// TwinCAT 3 PLC project MainControl
// ProgramVersion: 3.1.4024.0
// libraries:
//   JS_MC_REF, * (Jenny Science AG)
//   Tc2_EtherCAT, * (Beckhoff Automation GmbH)
//   Tc2_MC2, * (Beckhoff Automation GmbH)
//   Tc2_NCI, * (Beckhoff Automation GmbH)
//   Tc2_PlcInterpolation, * (Beckhoff Automation GmbH)
//   Tc2_Standard, * (Beckhoff Automation GmbH)
//   Tc2_System, * (Beckhoff Automation GmbH)
//   Tc2_Utilities, * (Beckhoff Automation GmbH)
//   Tc3_Module, * (Beckhoff Automation GmbH)
// project tree:
//   DUTs/ MFuncs.TcDUT, T_StringQueue.TcDUT
//   GVLs/ ExtPort.TcGVL, HMIVar.TcGVL, PYADSPort.TcGVL, UserVar.TcGVL
//   / PlcTask.TcTTO
//   POUs/FB/ FB_BackendManager.TcPOU, FB_ExtMessage.TcPOU, FB_HMITask.TcPOU, FB_JSReference.TcPOU, FB_Jog.TcPOU, FB_McodeMonitor.TcPOU, FB_MotorPower.TcPOU, FB_MotorReset.TcPOU, FB_RParamInit.TcPOU, FB_TimeCalculator.TcPOU
//   POUs/FB/Keyence/ FB_LJ_S8000Capture.TcPOU
//   POUs/FB/MicroFab/ FB_PulseInterval.TcPOU
//   POUs/FB/Nordson/ FB_ReadPressure.TcPOU, FB_WritePressure.TcPOU
//   POUs/function/ f_Contains_INT.TcPOU, f_MakeAbsPath.TcPOU, f_QueuePop.TcPOU, f_QueuePush.TcPOU, f_Queue_ToString.TcPOU
//   POUs/ MotorControl.TcPOU
// real-time tasks:
//   TASK PlcTask: cycle T#10ms, priority 20, ADS port 350
// motion (NC):
//   TASK NC-Task 1 SAF: cycle T#1ms, priority 4, ADS port 501
//   TASK NC-Task 1 SVB: cycle T#10ms, priority 8, ADS port 511
//   AXIS Axis 1 (id 1)
//     Velo: SlowManual=5, FastManual=30, Maximum=4500
//     OtherSettings: AllowMotionCmdToSlave=true
//     encoder EncType=19
//       EncPara: ScaleFactorNumerator=0.001, MaxCount=#xffffffff
//     drive DrvType=16
//       DrvPara: MaxCount=#xffffffff, DriveControlDWord=#x00020100
//         Analog: VeloReferenz=4500, VeloScale=125, AccScale=0.02, TorqueSetpointScale=10, ScaleFactorActTorque=0.1
//         TimeComp: TaskDelayCycles=1
//     controller CtrType=9
//       CtrPara: PriorControlFactor=1
//         Observer: BandWidth=20
//   AXIS Axis 2 (id 2)
//     Velo: SlowManual=5, FastManual=30, Maximum=4500
//     OtherSettings: AllowMotionCmdToSlave=true
//     encoder EncType=19
//       EncPara: ScaleFactorNumerator=0.001, MaxCount=#xffffffff
//     drive DrvType=16
//       DrvPara: MaxCount=#xffffffff, DriveControlDWord=#x00020100
//         Analog: VeloReferenz=4500, VeloScale=125, AccScale=0.02, TorqueSetpointScale=10, ScaleFactorActTorque=0.1
//         TimeComp: TaskDelayCycles=1
//     controller CtrType=9
//       CtrPara: PriorControlFactor=1
//         PID: PosKp=0
//         Observer: BandWidth=20
//   AXIS Axis 3 (id 3)
//     Velo: SlowManual=5, FastManual=30, Maximum=4500
//     OtherSettings: AllowMotionCmdToSlave=true
//     encoder EncType=19
//       EncPara: ScaleFactorNumerator=0.001, MaxCount=#xffffffff
//     drive DrvType=16
//       DrvPara: MaxCount=#xffffffff, DriveControlDWord=#x00020100
//         Analog: VeloReferenz=4500, VeloScale=125, AccScale=0.02, TorqueSetpointScale=10, ScaleFactorActTorque=0.1
//         TimeComp: TaskDelayCycles=1
//     controller CtrType=9
//       CtrPara: PriorControlFactor=1
//         Observer: BandWidth=20
//   AXIS Axis 4 (id 4)
//     Velo: SlowManual=1, FastManual=5
//     OtherSettings: AllowMotionCmdToSlave=true
//     encoder EncType=19
//       EncPara: MaxCount=#xffffffff
//     drive DrvType=16
//       DrvPara: MaxCount=#xffffffff, DriveControlDWord=#x00020000
//         Analog: TorqueSetpointScale=10, ScaleFactorActTorque=0.1
//         TimeComp: TaskDelayCycles=1
//     controller CtrType=1
//       CtrPara: PriorControlFactor=1
//         Observer: BandWidth=20
// I/O:
//   DEVICE Device 2 (EtherCAT), AmsNetId 192.168.0.2.3.1
//     Drive 1 (Xvi) [XENAX Xvi 75V8S]
//     Drive 2 (Xvi) [XENAX Xvi 75V8S]
//     Drive 3 (Xvi) [XENAX Xvi 75V8S]
//     Drive 12 (Ezi-SERVO2 EtherCAT) [Ezi-SERVO2 EtherCAT]
//     Term 4 (EK1100) [EK1100 EtherCAT Coupler (2A E-Bus)]
//       Term 5 (EL1008) [EL1008 8Ch. Dig. Input 24V, 3ms]
//       Term 17 (EL2008) [EL2008 8Ch. Dig. Output 24V, 0.5A]
//       Term 6 (EL9185) [EL9185 Potential Connection, 4 x 24-230V]
//       Term 7 (EL9505) [EL9505 Power supply terminal 5V]
//       Term 10 (EL2124) [EL2124 4Ch. Dig. Output 5V, 20mA]
//       Term 11 (EL2634) [EL2634 4Ch. Relay Output, NO (250V AC / 30V DC)]
//       Term 9 (EL9011) [EL9011 End Terminal]
//     Box 8 (LJ-S_CB-NEC Series) [LJ-S_CB-NEC Series]
//       modules: Module 1 (Result Data 128Byte), Module 2 (Parameter 128Byte)
// variable links:
//   NC-Task 1 SAF/Axes/Axis 1 <-> Device 2 (EtherCAT)/Drive 1 (Xvi)
//     Drive/Inputs/In/nDataIn1 <-> 1. TxPDO CSP/Following Error Actual Value
//     Drive/Inputs/In/nState1 <-> 1. TxPDO CSP/Statusword
//     Drive/Inputs/In/nState2 <-> 1. TxPDO CSP/Statusword @bit 8
//     Drive/Inputs/In/nState4 @bit 1 <-> WcState/InputToggle
//     Drive/Inputs/In/nState4 <-> WcState/WcState
//     Drive/Outputs/Out/nCtrl1 <-> 1. RxPDO CSP/Controlword
//     Drive/Outputs/Out/nCtrl2 <-> 1. RxPDO CSP/Controlword @bit 8
//     Drive/Outputs/Out/nDataOut1 <-> 1. RxPDO CSP/Target Position
//     Drive/Outputs/Out/nDataOut2 <-> 4. RxPDO CSP FeedForward/Target Velocity
//     Drive/Outputs/Out/nDataOut3[0] <-> 4. RxPDO CSP FeedForward/Torque Offset
//     Enc/Inputs/In/nDataIn1 <-> 1. TxPDO CSP/Position Actual Value
//     Enc/Inputs/In/nState4 @bit 1 <-> WcState/InputToggle
//     Enc/Inputs/In/nState4 <-> WcState/WcState
//   NC-Task 1 SAF/Axes/Axis 2 <-> Device 2 (EtherCAT)/Drive 2 (Xvi)
//     Drive/Inputs/In/nDataIn1 <-> 1. TxPDO CSP/Following Error Actual Value
//     Drive/Inputs/In/nState1 <-> 1. TxPDO CSP/Statusword
//     Drive/Inputs/In/nState2 <-> 1. TxPDO CSP/Statusword @bit 8
//     Drive/Inputs/In/nState4 @bit 1 <-> WcState/InputToggle
//     Drive/Inputs/In/nState4 <-> WcState/WcState
//     Drive/Outputs/Out/nCtrl1 <-> 1. RxPDO CSP/Controlword
//     Drive/Outputs/Out/nCtrl2 <-> 1. RxPDO CSP/Controlword @bit 8
//     Drive/Outputs/Out/nDataOut1 <-> 1. RxPDO CSP/Target Position
//     Drive/Outputs/Out/nDataOut2 <-> 4. RxPDO CSP FeedForward/Target Velocity
//     Drive/Outputs/Out/nDataOut3[0] <-> 4. RxPDO CSP FeedForward/Torque Offset
//     Enc/Inputs/In/nDataIn1 <-> 1. TxPDO CSP/Position Actual Value
//     Enc/Inputs/In/nState4 @bit 1 <-> WcState/InputToggle
//     Enc/Inputs/In/nState4 <-> WcState/WcState
//   NC-Task 1 SAF/Axes/Axis 3 <-> Device 2 (EtherCAT)/Drive 3 (Xvi)
//     Drive/Inputs/In/nDataIn1 <-> 1. TxPDO CSP/Following Error Actual Value
//     Drive/Inputs/In/nState1 <-> 1. TxPDO CSP/Statusword
//     Drive/Inputs/In/nState2 <-> 1. TxPDO CSP/Statusword @bit 8
//     Drive/Inputs/In/nState4 @bit 1 <-> WcState/InputToggle
//     Drive/Inputs/In/nState4 <-> WcState/WcState
//     Drive/Outputs/Out/nCtrl1 <-> 1. RxPDO CSP/Controlword
//     Drive/Outputs/Out/nCtrl2 <-> 1. RxPDO CSP/Controlword @bit 8
//     Drive/Outputs/Out/nDataOut1 <-> 1. RxPDO CSP/Target Position
//     Drive/Outputs/Out/nDataOut2 <-> 4. RxPDO CSP FeedForward/Target Velocity
//     Drive/Outputs/Out/nDataOut3[0] <-> 4. RxPDO CSP FeedForward/Torque Offset
//     Enc/Inputs/In/nDataIn1 <-> 1. TxPDO CSP/Position Actual Value
//     Enc/Inputs/In/nState4 @bit 1 <-> WcState/InputToggle
//     Enc/Inputs/In/nState4 <-> WcState/WcState
//   NC-Task 1 SAF/Axes/Axis 4 <-> Device 2 (EtherCAT)/Drive 12 (Ezi-SERVO2 EtherCAT)
//     Drive/Inputs/In/nDcOutputTime <-> InfoData/DcOutputShift
//     Drive/Inputs/In/nState1 <-> CSP Inputs/Status Word
//     Drive/Inputs/In/nState2 <-> CSP Inputs/Status Word @bit 8
//     Drive/Inputs/In/nState4 @bit 1 <-> WcState/InputToggle
//     Drive/Inputs/In/nState4 <-> WcState/WcState
//     Drive/Outputs/Out/nCtrl1 <-> CSP Outputs/Control Word
//     Drive/Outputs/Out/nCtrl2 <-> CSP Outputs/Control Word @bit 8
//     Drive/Outputs/Out/nDataOut1 <-> CSP Outputs/Target Position
//     Enc/Inputs/In/nDataIn1 <-> CSP Inputs/Position Actual Value
//     Enc/Inputs/In/nDataIn3 <-> CSP Inputs/Touch probe 1 positive value
//     Enc/Inputs/In/nDataIn5 <-> CSP Inputs/Touch probe 2 positive value
//     Enc/Inputs/In/nDcInputTime <-> InfoData/DcInputShift
//     Enc/Inputs/In/nState4 @bit 1 <-> WcState/InputToggle
//     Enc/Inputs/In/nState4 <-> WcState/WcState
//     Enc/Inputs/In/nState5 <-> CSP Inputs/Touch probe status
//     Enc/Inputs/In/nState6 <-> CSP Inputs/Touch probe status @bit 8
//     Enc/Outputs/Out/nCtrl5 <-> CSP Outputs/Touch probe function
//     Enc/Outputs/Out/nCtrl6 <-> CSP Outputs/Touch probe function @bit 8
//   MainControl/MainControl Instance <-> Device 2 (EtherCAT)/Box 8 (LJ-S_CB-NEC Series)
//     PlcTask Inputs/ExtPort.LJ_S8000_bBusy <-> StatusBit/BUSY
//     PlcTask Inputs/ExtPort.LJ_S8000_bReady <-> StatusBit/READY
//     PlcTask Inputs/ExtPort.LJ_S8000_bTRG_ack <-> StatusBit/TRG_ack
//     PlcTask Outputs/ExtPort.LJ_S8000_bTRG <-> ControlBit/TRG
//   MainControl/MainControl Instance <-> Device 2 (EtherCAT)/Drive 1 (Xvi)
//     PlcTask Inputs/MotorControl.fb_JSReference.JS_MC_X.stSlaveAmsAddr <-> InfoData/AdsAddr
//   MainControl/MainControl Instance <-> Device 2 (EtherCAT)/Drive 2 (Xvi)
//     PlcTask Inputs/MotorControl.fb_JSReference.JS_MC_Y.stSlaveAmsAddr <-> InfoData/AdsAddr
//   MainControl/MainControl Instance <-> Device 2 (EtherCAT)/Drive 3 (Xvi)
//     PlcTask Inputs/MotorControl.fb_JSReference.JS_MC_Z.stSlaveAmsAddr <-> InfoData/AdsAddr
//   MainControl/MainControl Instance <-> Device 2 (EtherCAT)/Term 4 (EK1100)/Term 10 (EL2124)
//     PlcTask Outputs/ExtPort.EL2124_OUT[0] <-> Channel 1/Output
//   MainControl/MainControl Instance <-> Device 2 (EtherCAT)/Term 4 (EK1100)/Term 11 (EL2634)
//     PlcTask Outputs/ExtPort.EL2634_OUT[0] <-> Channel 1/Output
//   MainControl/MainControl Instance <-> Device 2 (EtherCAT)/Term 4 (EK1100)/Term 5 (EL1008)
//     PlcTask Inputs/ExtPort.EL1008_IN[0] <-> Channel 1/Input
//     PlcTask Inputs/ExtPort.EL1008_IN[1] <-> Channel 2/Input
//   MainControl/MainControl Instance <-> NC-Task 1 SAF/Axes/Axis 1
//     PlcTask Inputs/MotorControl.motX.NcToPlc <-> Outputs/ToPlc
//     PlcTask Outputs/MotorControl.motX.PlcToNc <-> Inputs/FromPlc
//   MainControl/MainControl Instance <-> NC-Task 1 SAF/Axes/Axis 2
//     PlcTask Inputs/MotorControl.motY.NcToPlc <-> Outputs/ToPlc
//     PlcTask Outputs/MotorControl.motY.PlcToNc <-> Inputs/FromPlc
//   MainControl/MainControl Instance <-> NC-Task 1 SAF/Axes/Axis 3
//     PlcTask Inputs/MotorControl.motZ.NcToPlc <-> Outputs/ToPlc
//     PlcTask Outputs/MotorControl.motZ.PlcToNc <-> Inputs/FromPlc
//   MainControl/MainControl Instance <-> NC-Task 1 SAF/Axes/Axis 4
//     PlcTask Inputs/MotorControl.motQ1.NcToPlc <-> Outputs/ToPlc
//     PlcTask Outputs/MotorControl.motQ1.PlcToNc <-> Inputs/FromPlc
//   MainControl/MainControl Instance <-> NC-Task 1 SAF/Channel 2
//     PlcTask Inputs/MotorControl.inst_NcToPlc_NCI <-> Outputs/ToPlc
//     PlcTask Outputs/MotorControl.inst_PlcToNc_NCI <-> Inputs/FromPlc

CONFIGURATION MainControl
    RESOURCE PLC ON TwinCAT3
        TASK PlcTask(INTERVAL := T#10ms, PRIORITY := 20);
        PROGRAM MotorControl WITH PlcTask : MotorControl;
    END_RESOURCE
END_CONFIGURATION

// ---- DUTs/MFuncs.TcDUT
TYPE MFuncs :
//	M: 0 ~ 159
//	NOT TO USE THESE M-FUNCTIONS
//  2	(Program end)
//	17	(End of subprogram)
//	30	(Program end with delection of all fast M functions)
(
	M_NordsonExtOn		:=	10,
	M_NordsonExtOff 	:=	11,

	M_MicrofabExtOn		:=	20,
	M_MicrofabExtOff	:=	21,
	
	M_LJ_S8000TRG		:=	50,
	
	
	M_NordsonPresTRG100	:=	100,
	M_NordsonPresTRG101	:=	101,
	M_NordsonPresTRG102	:=	102,
	M_NordsonPresTRG103	:=	103,
	M_NordsonPresTRG104	:=	104,
	M_NordsonPresTRG105	:=	105,
	M_NordsonPresTRG106	:=	106,
	M_NordsonPresTRG107	:=	107,
	M_NordsonPresTRG108	:=	108,
	M_NordsonPresTRG109	:=	109,
	
	M_MicrofabIntTRG110 :=	110,
	M_MicrofabIntTRG111 :=	111,
	M_MicrofabIntTRG112 :=	112,
	
	
	M_RHskTRG			:=	150
	
);
END_TYPE

// ---- DUTs/T_StringQueue.TcDUT
TYPE T_StringQueue :
STRUCT
    Buffer : ARRAY[0..19] OF STRING(255); // 큐 크기 20
    Head   : INT	:=	0;  // Pop 위치
    Tail   : INT	:=	0;  // Push 위치
    Count  : INT	:=	0;  // 현재 개수
END_STRUCT
END_TYPE

// ---- GVLs/ExtPort.TcGVL
{attribute 'qualified_only'}
VAR_GLOBAL
	// ExtPort.EL2124_OUT[0]	:	MicroFab Ext 1
	EL2124_OUT	AT%Q*	:	ARRAY[0..3]	OF	BOOL;
	
	// ExtPort.EL2634_OUT[0]	:	Nordson Ext 1
	EL2634_OUT	AT%Q*	:	ARRAY[0..3]	OF	BOOL;
	
	LJ_S8000_bBusy		AT%I*	:	BOOL;
	LJ_S8000_bTRG_ack	AT%I*	:	BOOL;
	LJ_S8000_bReady		AT%I*	:	BOOL;
	LJ_S8000_bTRG		AT%Q*	:	BOOL;
	
	EL1008_IN	AT%I*	:	ARRAY[0..7]	OF	BOOL;
END_VAR

// ---- GVLs/HMIVar.TcGVL
{attribute 'qualified_only'}
VAR_GLOBAL
	
	sActPosX	:	STRING(32)	:=	'0.000';
	sActPosY	:	STRING(32)	:=	'0.000';
	sActPosZ	:	STRING(32)	:=	'0.000';
	
	sActVelX	:	STRING(32)	:=	'0.000';
	sActVelY	:	STRING(32)	:=	'0.000';
	sActVelZ	:	STRING(32)	:=	'0.000';
	
	sActAccX	:	STRING(32)	:=	'0.000';
	sActAccY	:	STRING(32)	:=	'0.000';
	sActAccZ	:	STRING(32)	:=	'0.000';
	
	sSetPosX	:	STRING(32)	:=	'0.000';
	sSetPosY	:	STRING(32)	:=	'0.000';
	sSetPosZ	:	STRING(32)	:=	'0.000';
	
	sSetVelX	:	STRING(32)	:=	'0.000';
	sSetVelY	:	STRING(32)	:=	'0.000';
	sSetVelZ	:	STRING(32)	:=	'0.000';
	
	sSetAccX	:	STRING(32)	:=	'0.000';
	sSetAccY	:	STRING(32)	:=	'0.000';
	sSetAccZ	:	STRING(32)	:=	'0.000';
	
	
	EstimatedTime		:	STRING(32)	:=	'0.000s';
	
	
	bNaviActive	:	BOOL	:=	TRUE;
	
	CodeName	:	STRING(255);
	
	GCodeQueueString:	STRING(8192):=	'';
	
	NordsonPressure			:	STRING	:=	'0';
	
	
	I_ForceActX		AT%I*	:	DINT;
	I_ForceActY		AT%I*	:	DINT;
	I_ForceActZ		AT%I*	:	DINT;
	
	
	RunningGCodeLine	:	STRING(1024)	:=	'';
	
	CurrBlockNumSTR		:	STRING	:=	'-';
	
	
	
END_VAR

// ---- GVLs/PYADSPort.TcGVL
{attribute 'qualified_only'}
VAR_GLOBAL
	// Nordson
	bNordWriteReq	:	BOOL	:=	FALSE;
	bNordWriteErr	:	BOOL	:=	FALSE;
	bNordReadReq	:	BOOL	:=	FALSE;
	bNordReadErr	:	BOOL	:=	FALSE;
	nNordPress		:	REAL	:=	0.0;
	
	
	bHeartbeat		:	BOOL	:=	FALSE;
	dtHeartbeatTime	:	DT;
	
	bEstTimeReq		:	BOOL	:=	FALSE;
	bEstTimeErr		:	BOOL	:=	FALSE;
	nEstTime		:	REAL	:=	0.0;	
	
END_VAR

// ---- GVLs/UserVar.TcGVL
{attribute 'qualified_only'}
VAR_GLOBAL
	
	RunningGCodeName:	STRING(255)	:=	'';
//	QueuedGCodeName	:	STRING(255)	:=	'';
	GCodeNameQueue	:	T_StringQueue;
	
	ContinueGCode	:	BOOL	:=	TRUE;
	
	SingleGCodeMode	:	BOOL	:=	FALSE;
	SingleGCodeTRG	:	BOOL	:=	FALSE;
	
	// 0: OFF, 1: JOG, 2: GCODE
	OpMode	:	UDINT	:=	0;
	
	// 0: Nothing, +1: +, +2: ++, -1: -, -2: --
	// +-3: ManualVel 
	JogButtonX	:	INT	:=	0;
	JogButtonY	:	INT	:=	0;
	JogButtonZ	:	INT	:=	0;
//	JogVel		:	LREAL	:=	30.0;
	
	JogMovePos	:	BOOL	:=	FALSE;
	JogTargX	:	STRING	:=	'100.0';
	JogTargY	:	STRING	:=	'260.0';
	JogTargZ	:	STRING	:=	'60.0';
	JogTargVel	:	STRING	:=	'1800'; // Feedrate (mm/min)
	
	JogPowerX	:	BOOL	:=	TRUE;
	JogPowerY	:	BOOL	:=	TRUE;
	JogPowerZ	:	BOOL	:=	TRUE;
	
	NordsonReadPressureBtn	:	BOOL	:=	FALSE;
	NordsonWritePressureBtn	:	BOOL	:=	FALSE;
	NordsonPressureActive	:	BOOL	:=	TRUE;
	
	LJ_S8000CaptureBtn		:	BOOL	:=	FALSE;
	LJ_S8000CaptureActive	:	BOOL	:=	TRUE;
	
	GCodeBasePath	:	STRING(255)	:=	'C:\\Users\\Administrator\\Desktop\\GCodes';

	// 0: Don't input HMIVar.CodeName into execution
	// 1: HMIVar.CodeName into QueuedGCodeName
	// 2: HMIVar.CodeName into GCodeName LIST
	Auto_CodeType	:	INT	:=	1;
	
	R_Params		:	ARRAY[0..12] OF INT	:=
						[100, 101, 102, 103, 104, 105, 106, 107, 108, 109,
						 110, 111, 112];
	
	R_InitVal		:	LREAL	:=	-1.0;
	
	bBackendStarted	:	BOOL	:=	FALSE;
	
	//	gDtFromPy : DT;      // Python이 써주는 시간(권장: UTC epoch seconds로 써서 DT에 저장)
//    gPlcNowDt : DT;      // PLC 로컬 현재시간을 DT로 변환해 저장(옵션)
    gDiffSec  : LINT;    // (PLC - Python) 차이[초]
    gInSync   : BOOL	:=	TRUE;    // 동기 여부
	gPlcStr: STRING(24);
    gPyStr    : STRING(24);
	
	bClearQueue	:	BOOL	:=	FALSE;
	
	
	bESTOP		:	BOOL	:=	FALSE;
	bRESET		:	BOOL	:=	FALSE;
	
	
	bSingleBlockMode	:	BOOL	:=	FALSE;
	
	bNordsonFoot	:	BOOL	:=	FALSE;
	
	CurrBlockNum		:	UDINT	:=	0;
	// Optional Axis 4. Non-retained; all motion permissions default OFF.
	Q1Commissioned : BOOL := FALSE; // Operator confirmation; NOT a safety function
	Q1Enable : BOOL := FALSE;
	Q1UseInGCode : BOOL := FALSE; // Sampled in state 200, held for whole queue run
	Q1Reset : BOOL := FALSE; // Rising edge, idle only
	Q1JogButton : INT := 0; // -1 / 0 / +1 only
	Q1JogVelocity : LREAL := 0.0; // NC units/second; validate before setting
END_VAR

// ---- POUs/MotorControl.TcPOU
PROGRAM MotorControl
VAR
	motX	:	AXIS_REF;
	motY	:	AXIS_REF;
	motZ	:	AXIS_REF;
	
	inst_NcToPlc_NCI	AT %I*	:	NCTOPLC_NCICHANNEL_REF;
	inst_PlcToNc_NCI	AT %Q*	:	PLCTONC_NCICHANNEL_REF;
	
	fb_JSReference	:	FB_JSReference;
	fb_MotorPower	:	FB_MotorPower;
	fb_MotorReset	:	FB_MotorReset;
	
	fb_McodeMonitor	:	FB_McodeMonitor;
	fb_RParamInit	:	FB_RParamInit;
	fb_Backend		:	FB_BackendManager;
	
	bPowered	:	BOOL;
	bMotorReset	:	BOOL;
	bError		:	BOOL;
	bBusy		:	BOOL;
	
	bOpMcodeMonitor	:	BOOL	:=	FALSE;
	
	nMotorControlState	:	UDINT	:= 0;
	nInterpreterState	:	UDINT	:= 0;
	nErrorState			:	UDINT;
	
	
	fb_BuildGroup	:	CfgBuild3DGroup;
	fb_LoadProgEx	:	ItpLoadProgEx;
	fb_StartStopEx	:	ItpStartStopEx;
	fb_ClearGroup	:	CfgReconfigGroup;
	fb_ResetEx		:	ItpResetEx2;
	
	fb_MCJogX		:	FB_Jog;
	fb_MCJogY		:	FB_Jog;
	fb_MCJogZ		:	FB_Jog;
	
	fb_MoveAbsX		:	MC_MoveAbsolute;
	fb_MoveAbsY		:	MC_MoveAbsolute;
	fb_MoveAbsZ		:	MC_MoveAbsolute;
	
	fb_ExtMessage	:	FB_ExtMessage;
	
	fb_HMITask		:	FB_HMITask;
	
//	nMoveAbsVel		:	REAL	:=	30.0;
	
	fb_MCHaltX		:	MC_Halt;
	fb_MCHaltY		:	MC_Halt;
	fb_MCHaltZ		:	MC_Halt;
	
	fb_ItpEStop		:	ItpEStopEx;
	
	// Axis 4 extension: link motQ1 to NC Axis 4 after PLC Rebuild.
	motQ1 : AXIS_REF;
	fb_Q1Power : MC_Power;
	fb_Q1Reset : MC_Reset;
	fb_Q1Jog : MC_Jog;
	fb_Q1Status : MC_ReadStatus;
	fb_Q1ResetEdge : R_TRIG;
	fb_BuildGroupQ1 : CfgBuildExt3DGroup;
	bQ1UseLatched : BOOL := FALSE;
	bQ1Reserved : BOOL := FALSE; // Conservative lock, cleared only after group removal
	bQ1Linked : BOOL;
	bQ1Enable : BOOL;
	bQ1ManualAllowed : BOOL;
	bQ1Ready : BOOL;
	bQ1BuildStarted : BOOL := FALSE;
	nQ1Interlock : UDINT := 0; // 0=none, 1=start not ready, 2=permission/power/mode lost
	fQ1ActPos : LREAL;
	fQ1ActVelo : LREAL;

END_VAR

// Axis 4 service. No writes to existing XYZ ready/power/reset signals.
bQ1Linked := motQ1.NcToPlc.AxisId = 4;
fb_Q1Status(Axis := motQ1, Enable := bQ1Linked);
IF UserVar.bESTOP THEN
	UserVar.Q1Enable := FALSE; // No automatic re-enable after ESTOP reset
	UserVar.Q1JogButton := 0;
END_IF
bQ1Enable := bQ1Linked AND UserVar.Q1Commissioned AND UserVar.Q1Enable
	AND NOT UserVar.bESTOP;
fb_Q1Power(Axis := motQ1, Enable := bQ1Enable,
	Enable_Positive := bQ1Enable, Enable_Negative := bQ1Enable, Override := 100.0);
bQ1ManualAllowed := NOT bQ1Reserved AND NOT UserVar.bESTOP
	AND ((nMotorControlState = 0) OR (nMotorControlState = 100));
fb_Q1ResetEdge(CLK := UserVar.Q1Reset);
fb_Q1Reset(Axis := motQ1,
	Execute := fb_Q1ResetEdge.Q AND bQ1Linked AND NOT bQ1Reserved
		AND NOT fb_Q1Jog.Busy AND NOT UserVar.bESTOP
		AND ((nMotorControlState = 0) OR (nMotorControlState = 100)
			OR (nMotorControlState = 200)));
fb_Q1Jog(Axis := motQ1, Mode := E_JogMode.MC_JOGMODE_CONTINOUS,
	Velocity := UserVar.Q1JogVelocity,
	JogForward := bQ1ManualAllowed AND bQ1Enable AND fb_Q1Power.Status
		AND NOT fb_Q1Reset.Busy AND NOT UserVar.Q1Reset
		AND (UserVar.Q1JogVelocity > 0.0) AND (UserVar.Q1JogButton = 1),
	JogBackwards := bQ1ManualAllowed AND bQ1Enable AND fb_Q1Power.Status
		AND NOT fb_Q1Reset.Busy AND NOT UserVar.Q1Reset
		AND (UserVar.Q1JogVelocity > 0.0) AND (UserVar.Q1JogButton = -1));
bQ1Ready := bQ1Enable AND fb_Q1Power.Status AND NOT fb_Q1Power.Error
	AND fb_Q1Status.Valid AND fb_Q1Status.StandStill AND NOT fb_Q1Status.Error
	AND NOT fb_Q1Status.ErrorStop AND NOT fb_Q1Jog.Busy AND NOT fb_Q1Jog.Error
	AND NOT fb_Q1Reset.Busy AND NOT fb_Q1Reset.Error AND NOT UserVar.Q1Reset
	AND (UserVar.Q1JogButton = 0);
fQ1ActPos := motQ1.NcToPlc.ActPos;
fQ1ActVelo := motQ1.NcToPlc.ActVelo;
IF (nMotorControlState = 200) AND NOT bQ1Reserved THEN
	bQ1UseLatched := UserVar.Q1UseInGCode;
	nQ1Interlock := 0;
END_IF
// A participating Q1 fault stops the shared channel; XYZ-only runs are unaffected.
IF bQ1Reserved AND (nMotorControlState >= 202) AND (nMotorControlState <= 261)
	AND (NOT bQ1Enable OR NOT fb_Q1Power.Status OR fb_Q1Power.Error
		OR NOT fb_Q1Status.Valid OR fb_Q1Status.Error OR fb_Q1Status.ErrorStop
		OR (UserVar.OpMode <> 2)) THEN
	nQ1Interlock := 2;
	nErrorState := nMotorControlState;
	bError := TRUE;
	nMotorControlState := 299;
END_IF

CASE nMotorControlState OF

0:
	// Mode Selecting
	IF (UserVar.OpMode = 1) OR (UserVar.OpMode = 2) THEN
		bBusy	:=	TRUE;
		nMotorControlState	:=	1;
	ELSE
		bBusy	:=	FALSE;
		bOpMcodeMonitor		:=	FALSE;
	END_IF

//1:
//	fb_MotorReset(
//		motX	:=	motX,
//		motY	:=	motY,
//		motZ	:=	motZ,
//		bResetX	:=	TRUE,
//		bResetY	:=	TRUE,
//		bResetZ	:=	TRUE,
//		bReset	=>	bMotorReset);
//	IF bMotorReset THEN
////		fb_MotorReset.bResetX	:=	FALSE;
////		fb_MotorReset.bResetY	:=	FALSE;
////		fb_MotorReset.bResetZ	:=	FALSE;
//		nMotorControlState	:= 2;
//	END_IF

1:
	// Initial Power ON
	fb_MotorPower(
		motX	:=	motX,
		motY	:=	motY,
		motZ	:=	motZ,
		bPowerX	:=	TRUE,
		bPowerY	:=	TRUE,
		bPowerZ	:=	TRUE,
		bPowered=>	bPowered);
	IF bPowered THEN
		nMotorControlState	:= 2;
	END_IF

2:
	// Initial Referencing
	fb_JSReference(
		motX	:=	motX,
		motY	:=	motY,
		motZ	:=	motZ,
		bStartX	:=	TRUE,
		bStartY	:=	TRUE,
		bStartZ	:=	TRUE);
	IF fb_JSReference.bReferenced THEN
		fb_JSReference.bStartX	:=	FALSE;
		fb_JSReference.bStartY	:=	FALSE;
		fb_JSReference.bStartZ	:=	FALSE;
		bBusy	:=	FALSE;
		IF UserVar.OpMode = 1 THEN
			nMotorControlState	:= 100;
		ELSIF UserVar.OpMode = 2 THEN
			nMotorControlState	:= 200;
		END_IF
	END_IF

50:
	fb_MotorPower(
		motX	:=	motX,
		motY	:=	motY,
		motZ	:=	motZ,
		bPowerX	:=	FALSE,
		bPowerY	:=	FALSE,
		bPowerZ	:=	FALSE);
	IF NOT fb_MotorPower.bPowerBusy THEN
		bBusy	:=	FALSE;
		nMotorControlState	:=	0;
	END_IF


90:
	UserVar.bRESET	:=	FALSE;
	nMotorControlState	:=	50;
	


99:
	IF UserVar.bRESET THEN
		UserVar.bESTOP	:=	FALSE;
		nMotorControlState	:=	90;
	END_IF
	

100:
	// Jog Mode
	IF 	(UserVar.JogButtonX <> 0) OR
		(UserVar.JogButtonY <> 0) OR
		(UserVar.JogButtonZ <> 0) THEN
		bBusy	:=	TRUE;
		nMotorControlState	:=	110;
	ELSIF UserVar.JogMovePos THEN
		bBusy	:=	TRUE;
		nMotorControlState	:=	120;
	ELSIF 	UserVar.NordsonReadPressureBtn OR
			UserVar.NordsonWritePressureBtn OR 
			UserVar.LJ_S8000CaptureBtn THEN
		bBusy	:=	TRUE;
		nMotorControlState	:=	130;	// HMI Task
	ELSE
		bBusy	:=	FALSE;
	END_IF
	
	IF	(fb_MotorPower.Power_X	<>	UserVar.JogPowerX) OR
		(fb_MotorPower.Power_Y	<>	UserVar.JogPowerY) OR
		(fb_MotorPower.Power_Z	<>	UserVar.JogPowerZ) THEN
		nMotorControlState	:=	101;
		bBusy	:=	TRUE;		
	END_IF
	
	IF UserVar.OpMode <> 1 THEN
		// Turning OFF
		bBusy	:=	TRUE;
		nMotorControlState	:=	50;
	END_IF

101:
	// Power Changed
	fb_MotorPower(
		motX	:=	motX,
		motY	:=	motY,
		motZ	:=	motZ,
		bPowerX	:=	UserVar.JogPowerX,
		bPowerY	:=	UserVar.JogPowerY,
		bPowerZ	:=	UserVar.JogPowerZ);
	IF NOT fb_MotorPower.bPowerBusy THEN
		fb_JSReference(
			motX	:=	motX,
			motY	:=	motY,
			motZ	:=	motZ,
			bStartX	:=	UserVar.JogPowerX,
			bStartY	:=	UserVar.JogPowerY,
			bStartZ	:=	UserVar.JogPowerZ);
		IF (NOT (UserVar.JogPowerX OR UserVar.JogPowerY OR UserVar.JogPowerZ))
			OR fb_JSReference.bReferenced THEN
			bBusy	:=	FALSE;
			nMotorControlState	:= 100;
		END_IF
	END_IF



	
	
110:
	fb_MCJogX(mot	:=	motX,
		JogButton	:=	BOOL_TO_INT(UserVar.JogPowerX) * UserVar.JogButtonX);
	fb_MCJogY(mot	:=	motY,
		JogButton	:=	BOOL_TO_INT(UserVar.JogPowerY) * UserVar.JogButtonY);
	fb_MCJogZ(mot	:=	motZ,
		JogButton	:=	BOOL_TO_INT(UserVar.JogPowerZ) * UserVar.JogButtonZ);

//	IF 
//	END_IF
	IF	(fb_MCJogX.bError OR 
		 fb_MCJogY.bError OR
		 fb_MCJogZ.bError) THEN
		nMotorControlState :=	199;
	ELSIF NOT (fb_MCJogX.bBusy OR
			fb_MCJogY.bBusy OR
			fb_MCJogZ.bBusy) THEN
		nMotorControlState	:=	100;
	END_IF

120:
	IF UserVar.JogPowerX THEN
		fb_MoveAbsX(
			Axis		:=	motX,
			position	:=	STRING_TO_LREAL(UserVar.JogTargX),
			velocity	:=	STRING_TO_LREAL(UserVar.JogTargVel)/60.0,
			Execute		:=	TRUE);
	END_IF
	IF UserVar.JogPowerY THEN
		fb_MoveAbsY(
			Axis		:=	motY,
			position	:=	STRING_TO_LREAL(UserVar.JogTargY),
			velocity	:=	STRING_TO_LREAL(UserVar.JogTargVel)/60.0,
			Execute		:=	TRUE);
	END_IF
	IF UserVar.JogPowerZ THEN
		fb_MoveAbsZ(
			Axis		:=	motZ,
			position	:=	STRING_TO_LREAL(UserVar.JogTargZ),
			velocity	:=	STRING_TO_LREAL(UserVar.JogTargVel)/60.0,
			Execute		:=	TRUE);
	END_IF
	nMotorControlState	:=	121;
	
	

121:
	IF UserVar.JogPowerX THEN
		fb_MoveAbsX(
			Axis		:=	motX,
			position	:=	STRING_TO_LREAL(UserVar.JogTargX),
			velocity	:=	STRING_TO_LREAL(UserVar.JogTargVel)/60.0,
			Execute		:=	FALSE);
	END_IF
	IF UserVar.JogPowerY THEN
		fb_MoveAbsY(
			Axis		:=	motY,
			position	:=	STRING_TO_LREAL(UserVar.JogTargY),
			velocity	:=	STRING_TO_LREAL(UserVar.JogTargVel)/60.0,
			Execute		:=	FALSE);
	END_IF
	IF UserVar.JogPowerZ THEN
		fb_MoveAbsZ(
			Axis		:=	motZ,
			position	:=	STRING_TO_LREAL(UserVar.JogTargZ),
			velocity	:=	STRING_TO_LREAL(UserVar.JogTargVel)/60.0,
			Execute		:=	FALSE);
	END_IF
	
	IF NOT ((UserVar.JogPowerX AND fb_MoveAbsX.Busy) OR
			(UserVar.JogPowerY AND fb_MoveAbsY.Busy) OR
			(UserVar.JogPowerZ AND fb_MoveAbsZ.Busy)) THEN
		UserVar.JogMovePos	:=	FALSE;
		bBusy	:=	FALSE;
		nMotorControlState	:=	100;
	END_IF

	
130:
	IF NOT (UserVar.NordsonReadPressureBtn OR
			UserVar.NordsonWritePressureBtn OR
			UserVar.LJ_S8000CaptureBtn) THEN
		bBusy	:=	FALSE;
		nMotorControlState	:= 100;
	END_IF


190:
	fb_MCHaltX(
		Axis	:=	motX,
		Execute	:=	FALSE);
	fb_MCHaltY(
		Axis	:=	motY,
		Execute	:=	FALSE);
	fb_MCHaltZ(
		Axis	:=	motZ,
		Execute	:=	FALSE);
	
	fb_MoveAbsX(
		Axis		:=	motX,
		Execute		:=	FALSE);
	fb_MoveAbsY(
		Axis		:=	motY,
		Execute		:=	FALSE);
	fb_MoveAbsZ(
		Axis		:=	motZ,
		Execute		:=	FALSE);
	
	nMotorControlState	:=	191;
		
191:	
	fb_MCJogX(mot	:=	motX,
		JogButton	:=	0);
	fb_MCJogY(mot	:=	motY,
		JogButton	:=	0);
	fb_MCJogZ(mot	:=	motZ,
		JogButton	:=	0);
	
	fb_MotorReset(
		motX	:=	motX,
		motY	:=	motY,
		motZ	:=	motZ,
		bResetX	:=	fb_MCJogX.bError,
		bResetY	:=	fb_MCJogY.bError,
		bResetZ	:=	fb_MCJogZ.bError,
		bReset	=>	bMotorReset);
		
	IF bMotorReset THEN
		nMotorControlState	:=	192;
	END_IF
	
	
192:
	fb_MotorReset(
		motX	:=	motX,
		motY	:=	motY,
		motZ	:=	motZ,
		bResetX	:=	FALSE,
		bResetY	:=	FALSE,
		bResetZ	:=	FALSE,
		bReset	=>	bMotorReset);

	nMotorControlState	:=	193;
	
193:
	fb_MCJogX(mot	:=	motX,
		JogButton	:=	0);
	fb_MCJogY(mot	:=	motY,
		JogButton	:=	0);
	fb_MCJogZ(mot	:=	motZ,
		JogButton	:=	0);
	
	UserVar.bRESET	:=	FALSE;
	UserVar.JogMovePos	:=	FALSE;
	nMotorControlState	:=	50;

	
199:
	fb_MCHaltX(
		Axis	:=	motX,
		Execute	:=	TRUE);
	fb_MCHaltY(
		Axis	:=	motY,
		Execute	:=	TRUE);
	fb_MCHaltZ(
		Axis	:=	motZ,
		Execute	:=	TRUE);
	IF (fb_MCHaltX.Done AND
		fb_MCHaltY.Done AND
		fb_MCHaltZ.Done)
		AND UserVar.bRESET THEN// AND bMotorReset THEN
		
		UserVar.bESTOP	:=	FALSE;
		nMotorControlState	:=	190;
	END_IF

	
	
200:
	IF UserVar.SingleGCodeMode THEN
		IF UserVar.SingleGCodeTRG THEN
			UserVar.SingleGCodeTRG	:=	FALSE;
			UserVar.RunningGCodeName	:=	HMIVar.CodeName;
			bBusy	:=	TRUE;
			bOpMcodeMonitor		:=	TRUE;
			nMotorControlState	:=	201;
		END_IF
	ELSE
		IF UserVar.ContinueGCode THEN
			IF f_QueuePop(
					pQueue := ADR(UserVar.GCodeNameQueue),
					str => UserVar.RunningGCodeName) THEN
				HMIVar.GCodeQueueString	:=	f_Queue_ToString(ADR(UserVar.GCodeNameQueue));
				bBusy	:=	TRUE;
				bOpMcodeMonitor		:=	TRUE;
				nMotorControlState	:=	201;
	//		ELSIF UserVar.OpMode <> 2 THEN
	//			// Turning OFF
	//			bBusy	:=	TRUE;
	//			nMotorControlState	:=	50;
			END_IF
	//	ELSIF UserVar.OpMode <> 2 THEN
	//		// Turning OFF
	//		bBusy	:=	TRUE;
	//		nMotorControlState	:=	50;
		END_IF
	END_IF

	IF UserVar.OpMode <> 2 THEN
		// Turning OFF
		bBusy	:=	TRUE;
		nMotorControlState	:=	50;
	END_IF

201:
	IF bQ1UseLatched THEN
		bQ1Reserved := TRUE;
		IF NOT bQ1BuildStarted AND NOT bQ1Ready THEN
			nQ1Interlock := 1;
			nErrorState := 201;
			bError := TRUE;
			nMotorControlState := 299;
		ELSE
	// Initial interpolation group building
	nInterpreterState	:=	ItpGetStateInterpreter(sNciToPlc:=inst_NcToPlc_NCI);
	IF	nInterpreterState = Tc2_NCI.NCI_INTERPRETER_IDLE	THEN	
		bQ1BuildStarted := TRUE;
		fb_BuildGroupQ1(
			bExecute	:= TRUE, 
			nGroupId	:= ItpGetGroupId(sNciToPlc:=inst_NcToPlc_NCI) , 
			nXAxisId	:= motX.NcToPlc.AxisId, 
			nYAxisId	:= motY.NcToPlc.AxisId, 
			nZAxisId	:= motZ.NcToPlc.AxisId,
			nQ1AxisId := motQ1.NcToPlc.AxisId,
			nQ2AxisId := 0, nQ3AxisId := 0, nQ4AxisId := 0, nQ5AxisId := 0);
		IF NOT fb_BuildGroupQ1.bBusy THEN
			IF NOT fb_BuildGroupQ1.bErr THEN
				fb_RParamInit(
					bExecute	:=	TRUE,
					inst_NcToPlc_NCI	:=	inst_NcToPlc_NCI);
				nMotorControlState	:= 202;
			ELSE
				nErrorState	:= nMotorControlState;
				bError	:= TRUE;
				nMotorControlState	:= 299;
			END_IF
			ItpSetOverridePercent(
				fOverridePercent	:=	100.0,
				sPlcToNci	:=	inst_PlcToNc_NCI);
		END_IF
	
	END_IF
		END_IF
	ELSE
	// Initial interpolation group building
	nInterpreterState	:=	ItpGetStateInterpreter(sNciToPlc:=inst_NcToPlc_NCI);
	IF	nInterpreterState = Tc2_NCI.NCI_INTERPRETER_IDLE	THEN	
		fb_BuildGroup(
			bExecute	:= TRUE, 
			nGroupId	:= ItpGetGroupId(sNciToPlc:=inst_NcToPlc_NCI) , 
			nXAxisId	:= motX.NcToPlc.AxisId, 
			nYAxisId	:= motY.NcToPlc.AxisId, 
			nZAxisId	:= motZ.NcToPlc.AxisId);
		IF NOT fb_BuildGroup.bBusy THEN
			IF NOT fb_BuildGroup.bErr THEN
				fb_RParamInit(
					bExecute	:=	TRUE,
					inst_NcToPlc_NCI	:=	inst_NcToPlc_NCI);
				nMotorControlState	:= 202;
			ELSE
				nErrorState	:= nMotorControlState;
				bError	:= TRUE;
				nMotorControlState	:= 299;
			END_IF
			ItpSetOverridePercent(
				fOverridePercent	:=	100.0,
				sPlcToNci	:=	inst_PlcToNc_NCI);
		END_IF
	
	END_IF
	END_IF

202:
	fb_BuildGroupQ1(bExecute := FALSE);
	fb_BuildGroup(	bExecute	:= FALSE	); 
	IF fb_RParamInit.bBusy THEN
		fb_RParamInit(
			bExecute	:=	FALSE,
			inst_NcToPlc_NCI	:=	inst_NcToPlc_NCI);
		nMotorControlState	:= 205;			
	END_IF

205:
	fb_RParamInit(
		bExecute	:=	FALSE,
		inst_NcToPlc_NCI	:=	inst_NcToPlc_NCI);
	IF NOT fb_RParamInit.bBusy THEN
		IF fb_RParamInit.bErr THEN
			nMotorControlState	:=	202;
		ELSE
			nMotorControlState	:=	210;
		END_IF
	END_IF
	

210:
	fb_LoadProgEx(
		sNciToPlc	:=	inst_NcToPlc_NCI,
		bExecute	:=	TRUE,
		sPrg		:=	f_MakeAbsPath(UserVar.RunningGCodeName),
		nLength		:=	INT_TO_UDINT(LEN(f_MakeAbsPath(UserVar.RunningGCodeName))));
	
	IF NOT fb_LoadProgEx.bBusy THEN
		IF NOT fb_LoadProgEx.bErr THEN
			nMotorControlState	:=	211;
		ELSE
			nErrorState	:=	nMotorControlState;
			bError	:=	TRUE;
			nMotorControlState	:=	299;
		END_IF
		fb_LoadProgEx(
			sNciToPlc	:=	inst_NcToPlc_NCI,
			bExecute	:=	FALSE); 
	END_IF
	
	
211:
	fb_StartStopEx(
		bStart	:=	TRUE,
		bStop	:=	FALSE,
		tTimeOut	:= , 
		sNciToPlc	:=	 inst_NcToPlc_NCI);
	
	IF NOT fb_StartStopEx.bBusy THEN
		IF NOT fb_StartStopEx.bErr THEN
			nMotorControlState	:=	212;
		ELSE
			nErrorState	:=	nMotorControlState;
			bError	:=	TRUE;
			nMotorControlState	:=	299;
		END_IF
		fb_StartStopEx(
			bStart	:=	FALSE,
			sNciToPlc	:=	 inst_NcToPlc_NCI); 
	END_IF
	
212:
	nInterpreterState	:= ItpGetStateInterpreter(sNciToPlc:=inst_NcToPlc_NCI);
	IF nInterpreterState <> Tc2_NCI.NCI_INTERPRETER_READY THEN
		// nci is running
		nMotorControlState	:= 213;
	END_IF


213:
	nInterpreterState	:= ItpGetStateInterpreter(sNciToPlc:=inst_NcToPlc_NCI);
	IF	nInterpreterState = Tc2_NCI.NCI_INTERPRETER_READY THEN
		// program has finished
		fb_RParamInit(
			bExecute	:=	TRUE,
			inst_NcToPlc_NCI	:=	inst_NcToPlc_NCI);
		nMotorControlState	:= 230;
	ELSIF 	nInterpreterState = Tc2_NCI.NCI_INTERPRETER_ABORTED 
	OR 		ItpHasError(sNciToPlc:=inst_NcToPlc_NCI)  THEN
		nErrorState	:= nMotorControlState;
		bError	:= TRUE;
		nMotorControlState	:= 299;
	END_IF
	
230:
	IF fb_RParamInit.bBusy THEN
		fb_RParamInit(
			bExecute	:=	FALSE,
			inst_NcToPlc_NCI	:=	inst_NcToPlc_NCI);
		nMotorControlState	:=	231;
	END_IF
	
231:
	fb_RParamInit(
		bExecute	:=	FALSE,
		inst_NcToPlc_NCI	:=	inst_NcToPlc_NCI);
	IF NOT fb_RParamInit.bBusy THEN
		IF fb_RParamInit.bErr THEN
			nMotorControlState	:=	213;
		ELSE
			nMotorControlState	:=	250;
		END_IF
	END_IF
	
250:
	IF (NOT UserVar.SingleGCodeMode) AND UserVar.ContinueGCode THEN
		IF f_QueuePop(
				pQueue := ADR(UserVar.GCodeNameQueue),
				str => UserVar.RunningGCodeName) THEN
			HMIVar.GCodeQueueString	:=	f_Queue_ToString(ADR(UserVar.GCodeNameQueue));
			nMotorControlState	:=	210;
		ELSE
			nMotorControlState	:=	260;
		END_IF
	ELSE
		nMotorControlState	:=	260;
	END_IF
	
260:
	fb_ClearGroup(
		bExecute	:= TRUE, 
		nGroupId	:= ItpGetGroupId(sNciToPlc:=inst_NcToPlc_NCI));

	IF NOT fb_ClearGroup.bBusy THEN
		IF NOT fb_ClearGroup.bErr THEN
			bQ1Reserved := FALSE;
			bQ1BuildStarted := FALSE;
			fb_BuildGroupQ1(bExecute := FALSE);
			nMotorControlState	:= 261;
		ELSE
			(* add error handling *)
			nErrorState	:= nMotorControlState;
			bError	:= TRUE;
			nMotorControlState	:= 299;				
		END_IF
		fb_ClearGroup(bExecute:=FALSE); 
	END_IF

261:
	fb_ResetEx(
		bExecute:= TRUE, 
		tTimeOut:= , 
		sNciToPlc:= inst_NcToPlc_NCI, 
		bBusy=> , 
		bErr=> , 
		nErrId=> );

	IF NOT fb_ResetEx.bBusy THEN
		IF NOT fb_ResetEx.bErr THEN
			bBusy	:=	FALSE;
			bOpMcodeMonitor		:=	FALSE;
			nMotorControlState	:=	200;
		ELSE
			(* add error handling *)
			nErrorState	:= nMotorControlState;
			bError	:= TRUE;
			nMotorControlState	:= 299;
		END_IF
		fb_ResetEx( bExecute:= FALSE, sNciToPlc:= inst_NcToPlc_NCI);
	END_IF

	
290:
	IF ItpIsEStopEx(inst_NcToPlc_NCI) THEN
		fb_ItpEStop(
			sNciToPlc	:=	inst_NcToPlc_NCI,
			bExecute	:=	FALSE);
		nMotorControlState	:=	291;
	END_IF

	
291:
	fb_ResetEx(
		bExecute:= TRUE, 
		sNciToPlc:= inst_NcToPlc_NCI);

	IF NOT fb_ResetEx.bBusy THEN
		IF NOT fb_ResetEx.bErr THEN
			bBusy	:=	FALSE;
			bOpMcodeMonitor		:=	FALSE;
			nMotorControlState	:=	292;
		ELSE
			nErrorState	:= nMotorControlState;
			bError	:= TRUE;
			nMotorControlState	:= 9999;
		END_IF
		fb_ResetEx( bExecute:= FALSE, sNciToPlc:= inst_NcToPlc_NCI);
	END_IF
	

292:
	fb_ClearGroup(
		bExecute	:= TRUE, 
		nGroupId	:= ItpGetGroupId(sNciToPlc:=inst_NcToPlc_NCI));

	IF NOT fb_ClearGroup.bBusy THEN
		IF NOT fb_ClearGroup.bErr THEN
			bQ1Reserved := FALSE;
			bQ1BuildStarted := FALSE;
			fb_BuildGroupQ1(bExecute := FALSE);
			nMotorControlState	:= 50;
		ELSE
			nErrorState	:= nMotorControlState;
			bError	:= TRUE;
			nMotorControlState	:= 9999;				
		END_IF
		fb_ClearGroup(bExecute:=FALSE); 
	END_IF


	
	
299:
	fb_ItpEStop(
		sNciToPlc	:=	inst_NcToPlc_NCI,
		bExecute	:=	TRUE);
	IF UserVar.bRESET THEN
		UserVar.ContinueGCode	:=	FALSE;
		UserVar.bClearQueue	:=	TRUE;
		UserVar.bESTOP	:=	FALSE;
		nMotorControlState	:=	290;
	END_IF

	
9999:
	// No Answer
	bBusy	:=	TRUE;

END_CASE




IF UserVar.bESTOP THEN
	// ESTOP button Triggered	-->	bESTOP: TRUE
	// ESTOP button released	-->	bESTOP: TRUE
	// RESET button Triggered	--> bRESET: TRUE, bESTOP: FALSE
		// 99/199/299 --> 90/190/290 (at eash state)
	// 9-/19-/29- --> 50	: bRESET: FALSE
	bBusy	:=	TRUE;
	CASE UserVar.OpMode OF
		0:
			nMotorControlState	:=	99;
		1:
			nMotorControlState	:=	199;
		2:
			nMotorControlState	:=	299;
	END_CASE
ELSE
	UserVar.bRESET	:=	FALSE;
END_IF






// Q1 reservation owns the NCI stop path even if OpMode was changed.
IF bQ1Reserved AND UserVar.bESTOP THEN
	nMotorControlState := 299;
END_IF

fb_HMITask();
fb_Backend();



(* CASE-INDEPENDENT LOOPS *)
fb_ExtMessage(
	inst_NcToPlc_NCI	:=	inst_NcToPlc_NCI,
	inst_PlcToNc_NCI	:=	inst_PlcToNc_NCI,
	motX	:=	motX,
	motY	:=	motY,
	motZ	:=	motZ,
	bBusy	:=	bBusy);

IF bOpMcodeMonitor	THEN
	fb_McodeMonitor(
		inst_NcToPlc_NCI	:=	inst_NcToPlc_NCI,
		inst_PlcToNc_NCI	:=	inst_PlcToNc_NCI);
END_IF

END_PROGRAM

// ---- POUs/FB/FB_JSReference.TcPOU
FUNCTION_BLOCK FB_JSReference
VAR_INPUT
	bStartX	:	BOOL;
	bStartY	:	BOOL;
	bStartZ	:	BOOL;
END_VAR
VAR_OUTPUT
	bReferenced: BOOL := FALSE;
END_VAR
VAR_IN_OUT
	motX:	AXIS_REF;
	motY:	AXIS_REF;
	motZ:	AXIS_REF;
END_VAR	
VAR
	JS_MC_X :	JS_MC_REF;
	JS_MC_Y :	JS_MC_REF;
	JS_MC_Z :	JS_MC_REF;
	Done_X	:	BOOL;
	Done_Y	:	BOOL;
	Done_Z	:	BOOL;
END_VAR

JS_MC_X(
	Axis	:=	motX,
	bExecute:=	bStartX,
	bAbort	:=	FALSE,
	bForceNewRef	:=FALSE,
	iTypeGantry	:=0,
	Done	=>	Done_X);
	
JS_MC_Y(
	Axis	:=	motY,
	bExecute:=	bStartY,
	bAbort	:=	FALSE,
	bForceNewRef	:=FALSE,
	iTypeGantry	:=0,
	Done	=>	Done_Y);
	
JS_MC_Z(
	Axis	:=	motZ,
	bExecute:=	bStartZ,
	bAbort	:=	FALSE,
	bForceNewRef	:=FALSE,
	iTypeGantry	:=0,
	Done	=>	Done_Z);

IF bStartX OR bStartY OR bStartZ THEN
	bReferenced	:=	
		((NOT bStartX) OR Done_X) AND
		((NOT bStartY) OR Done_Y) AND
		((NOT bStartZ) OR Done_Z);
ELSE
	bReferenced	:=	FALSE;
END_IF

END_FUNCTION_BLOCK

// ---- POUs/FB/FB_MotorPower.TcPOU
FUNCTION_BLOCK FB_MotorPower
VAR_INPUT
	bPowerX	:	BOOL;
	bPowerY	:	BOOL;
	bPowerZ	:	BOOL;
END_VAR
VAR_OUTPUT
	bPowered	:	BOOL	:=	FALSE;
	bPowerBusy	:	BOOL	:=	FALSE;	
	// Is valid even in POWER OFF operation
	// If axis is not off even if off operation input, then bPowered := FALSE
	
	Power_X	: 	BOOL;
	Power_Y	: 	BOOL;
	Power_Z	:	BOOL;
END_VAR
VAR_IN_OUT
	motX:	AXIS_REF;
	motY:	AXIS_REF;
	motZ:	AXIS_REF;
END_VAR	
VAR
	MC_POWER_X	:	MC_POWER;
	MC_POWER_Y	:	MC_POWER;
	MC_POWER_Z	:	MC_POWER;
	
	
END_VAR

MC_POWER_X(
	Axis	:=	motX,
	Enable	:=	bPowerX,
	Enable_Positive	:=	bPowerX,
	Enable_Negative	:=	bPowerX,
	Override:=	100.0,
	Status	=>	Power_X);

MC_POWER_Y(
	Axis	:=	motY,
	Enable	:=	bPowerY,
	Enable_Positive	:=	bPowerY,
	Enable_Negative	:=	bPowerY,
	Override:=	100.0,
	Status	=>	Power_Y);

MC_POWER_Z(
	Axis	:=	motZ,
	Enable	:=	bPowerZ,
	Enable_Positive	:=	bPowerZ,
	Enable_Negative	:=	bPowerZ,
	Override:=	100.0,
	Status	=>	Power_Z);


IF bPowerX OR bPowerY OR bPowerZ THEN
	bPowered	:=	
		((NOT bPowerX) OR Power_X) AND
		((NOT bPowerY) OR Power_Y) AND
		((NOT bPowerZ) OR Power_Z);
ELSE
	bPowered	:=	FALSE;
END_IF

bPowerBusy	:=
	(bPowerX XOR Power_X) OR
	(bPowerY XOR Power_Y) OR
	(bPowerZ XOR Power_Z);

END_FUNCTION_BLOCK

// ---- POUs/FB/FB_MotorReset.TcPOU
FUNCTION_BLOCK FB_MotorReset
VAR_INPUT
	bResetX	:	BOOL;
	bResetY	:	BOOL;
	bResetZ	:	BOOL;
END_VAR
VAR_OUTPUT
	bReset	: BOOL := FALSE;
END_VAR
VAR_IN_OUT
	motX:	AXIS_REF;
	motY:	AXIS_REF;
	motZ:	AXIS_REF;
END_VAR
VAR
	MC_RESET_X	:	MC_RESET;
	MC_RESET_Y	:	MC_RESET;
	MC_RESET_Z	:	MC_RESET;
	
	Done_X	:	BOOL;
	Done_Y	:	BOOL;
	Done_Z	:	BOOL;
END_VAR

MC_RESET_X(
	Axis	:=	motX,
	Execute	:=	bResetX,
	Done	=>	Done_X);
	
MC_RESET_Y(
	Axis	:=	motY,
	Execute	:=	bResetY,
	Done	=>	Done_Y);
	
MC_RESET_Z(
	Axis	:=	motZ,
	Execute	:=	bResetZ,
	Done	=>	Done_Z);
	
	
IF bResetX OR bResetY OR bResetZ THEN
	bReset	:=	
		((NOT bResetX) OR Done_X) AND
		((NOT bResetY) OR Done_Y) AND
		((NOT bResetZ) OR Done_Z);
ELSE
	bReset	:=	TRUE; ///
END_IF

END_FUNCTION_BLOCK

// ---- POUs/FB/FB_McodeMonitor.TcPOU
FUNCTION_BLOCK FB_McodeMonitor
VAR_INPUT
END_VAR
VAR_OUTPUT
END_VAR
VAR_IN_OUT
	inst_NcToPlc_NCI	:	NCTOPLC_NCICHANNEL_REF;
	inst_PlcToNc_NCI	:	PLCTONC_NCICHANNEL_REF;
END_VAR
VAR
	bNordsonExtOn		:	BOOL	:=	FALSE;
	bNordsonExtOff		:	BOOL	:=	FALSE;
	bMicrofabExtOn		:	BOOL	:=	FALSE;
	bMicrofabExtOff		:	BOOL	:=	FALSE;
	
	bLJ_S8000TRG		:	BOOL	:=	FALSE;
	nLJ_S8000State		:	UDINT	:=	0;
	
	bNordsonPresWriteTRG:	BOOL	:=	FALSE;	
	nNordsonPresWriteState	:	UDINT	:=	0;
	nNordsonPresRNum	:	INT	:=	0;	
	nNordsonPressRParam	:	LREAL	:=	0.0;
	
	nHskMNum			:	INT	:=	0;
	
	
	bRHskTRG			:	BOOL	:=	FALSE;
	nRHskState			:	UDINT	:=	0;
	nRHskBusyIdx			:	DINT	:=	0;
	nRHskVal			:	LREAL	:=	0;
	
	fb_ConfirmHsk		:	ItpConfirmHsk;
	fb_ReadRParams		:	ItpReadRParams;
	
	fb_LJ_S8000Cap		:	FB_LJ_S8000Capture;
	fb_WritePressure	:	FB_WritePressure;
	
	fb_MicroFabInterval	:	FB_PulseInterval;
	
	nMicroFabIntRNum	:	INT	:=	0;
	nMicroFabInterval	:	LREAL	:=	0.0;
	bMicroFabIntWriteTRG:	BOOL	:=	FALSE;
	nMicroFabIntWriteState	:	UDINT	:=	0;
	
END_VAR

bNordsonExtOn	:=	ItpIsFastMFunc(	
	nFastMFuncNo	:=	MFuncs.M_NordsonExtOn,
	sNciToPlc		:=	inst_NcToPlc_NCI);

bNordsonExtOff	:=	ItpIsFastMFunc(
	nFastMFuncNo	:=	MFuncs.M_NordsonExtOff,
	sNciToPlc		:=	inst_NcToPlc_NCI);

bMicrofabExtOn	:=	ItpIsFastMFunc(
	nFastMFuncNo	:=	MFuncs.M_MicrofabExtOn,
	sNciToPlc		:=	inst_NcToPlc_NCI);

bMicrofabExtOff	:=	ItpIsFastMFunc(
	nFastMFuncNo	:=	MFuncs.M_MicrofabExtOff,
	sNciToPlc		:=	inst_NcToPlc_NCI);

	

IF ItpIsHskMFunc(inst_NcToPlc_NCI) THEN
	nHskMNum	:=	ItpGetHskMFunc(inst_NcToPlc_NCI);
	IF f_Contains_INT(
		num	:=	nHskMNum,
		arr	:=	UserVar.R_Params) THEN
		IF (nHskMNum >= 100) AND (nHskMNum < 110) THEN
			nNordsonPresRNum		:=	nHskMNum;
			bNordsonPresWriteTRG	:=	TRUE;
		ELSIF (nHskMNum >= 110) AND (nHskMNum <= 112) THEN
			nMicroFabIntRNum		:=	nHskMNum;
			bMicroFabIntWriteTRG	:=	TRUE;
		END_IF
	ELSE
		CASE nHskMNum OF
			MFuncs.M_LJ_S8000TRG:
				bLJ_S8000TRG	:=	TRUE;
			MFuncs.M_RHskTRG:
				bRHskTRG	:=	TRUE;
		END_CASE
	END_IF
	
END_IF






IF bNordsonExtOn THEN
	ExtPort.EL2634_OUT[0] := TRUE;
ELSIF bNordsonExtOff THEN
	ExtPort.EL2634_OUT[0] := FALSE;
END_IF


IF bMicrofabExtOn THEN
	IF (nMicroFabInterval - 20) > -0.01 THEN
		fb_MicroFabInterval(
			bOn	:=	TRUE,
			nInterval	:=	TO_UDINT(nMicroFabInterval));
	ELSE
		fb_MicroFabInterval(
			bOn	:=	TRUE);
	END_IF
ELSIF bMicrofabExtOff THEN
	fb_MicroFabInterval(
		bOn	:=	FALSE);
END_IF
fb_MicroFabInterval();





IF bLJ_S8000TRG THEN
	CASE nLJ_S8000State	OF
		0:
			fb_LJ_S8000Cap(	bExecute	:=	TRUE);
			IF fb_LJ_S8000Cap.bBusy	THEN
				fb_LJ_S8000Cap.bExecute	:=	FALSE;
				nLJ_S8000State	:=	1;
			END_IF
		1:
			fb_LJ_S8000Cap(	bExecute	:=	FALSE);
			IF NOT fb_LJ_S8000Cap.bBusy THEN
				fb_ConfirmHsk(
					bExecute	:=	TRUE,
					sNciToPlc	:=	inst_NcToPlc_NCI,
					sPlcToNci	:=	inst_PlcToNc_NCI,);
				nLJ_S8000State	:=	2;
			END_IF
		2:
			IF 	fb_ConfirmHsk.bBusy THEN
				fb_ConfirmHsk(
					bExecute	:=	FALSE,
					sNciToPlc	:=	inst_NcToPlc_NCI,
					sPlcToNci	:=	inst_PlcToNc_NCI,);
				bLJ_S8000TRG	:=	FALSE;
				nLJ_S8000State	:=	0;
			END_IF
	END_CASE
END_IF



IF bNordsonPresWriteTRG THEN
	CASE nNordsonPresWriteState	OF
		0:
			fb_ReadRParams(
				bExecute	:=	TRUE,
				nChnId		:=	inst_NcToPlc_NCI.ChnId,
				pAddr		:=	ADR(nNordsonPressRParam),
				nIndex		:=	nNordsonPresRNum,
				nCount		:=	1);
			nNordsonPresWriteState	:=	1;
		1:
			IF fb_ReadRParams.bBusy THEN
				fb_ReadRParams(
					bExecute	:=	FALSE,
					nChnId		:=	inst_NcToPlc_NCI.ChnId,
					pAddr		:=	ADR(nNordsonPressRParam),
					nIndex		:=	nNordsonPresRNum,
					nCount		:=	1);
				fb_WritePressure(
					bExecute	:=	TRUE,
					Pressure	:=	LREAL_TO_REAL(nNordsonPressRParam));
				IF fb_WritePressure.bBusy	THEN
					nNordsonPresRNum	:=	0;
					fb_WritePressure.bExecute	:=	FALSE;
					nNordsonPresWriteState	:=	2;
				END_IF
			END_IF
		2:
			fb_WritePressure(	bExecute	:=	FALSE);
			IF NOT fb_WritePressure.bBusy THEN
				IF NOT fb_WritePressure.bErr THEN
					fb_ConfirmHsk(
						bExecute	:=	TRUE,
						sNciToPlc	:=	inst_NcToPlc_NCI,
						sPlcToNci	:=	inst_PlcToNc_NCI,);
					nNordsonPresWriteState	:=	3;
				ELSE
					nNordsonPresWriteState	:=	1;
				END_IF
			END_IF
		3:
			IF 	fb_ConfirmHsk.bBusy THEN
				fb_ConfirmHsk(
					bExecute	:=	FALSE,
					sNciToPlc	:=	inst_NcToPlc_NCI,
					sPlcToNci	:=	inst_PlcToNc_NCI,);
				bNordsonPresWriteTRG	:=	FALSE;
				nNordsonPresWriteState	:=	0;
			END_IF
	END_CASE
END_IF



IF bMicroFabIntWriteTRG THEN
	CASE nMicroFabIntWriteState	OF
		0:
			fb_ReadRParams(
				bExecute	:=	TRUE,
				nChnId		:=	inst_NcToPlc_NCI.ChnId,
				pAddr		:=	ADR(nMicroFabInterval),
				nIndex		:=	nMicroFabIntRNum,
				nCount		:=	1);
			nMicroFabIntWriteState	:=	1;
		1:
			IF fb_ReadRParams.bBusy THEN
				fb_ReadRParams(
					bExecute	:=	FALSE,
					nChnId		:=	inst_NcToPlc_NCI.ChnId,
					pAddr		:=	ADR(nMicroFabInterval),
					nIndex		:=	nMicroFabIntRNum,
					nCount		:=	1);
				fb_ConfirmHsk(
					bExecute	:=	TRUE,
					sNciToPlc	:=	inst_NcToPlc_NCI,
					sPlcToNci	:=	inst_PlcToNc_NCI,);
				nMicroFabIntWriteState	:=	2;
			END_IF
		2:
			IF 	fb_ConfirmHsk.bBusy THEN
				fb_ConfirmHsk(
					bExecute	:=	FALSE,
					sNciToPlc	:=	inst_NcToPlc_NCI,
					sPlcToNci	:=	inst_PlcToNc_NCI,);
				bMicroFabIntWriteTRG	:=	FALSE;
				nMicroFabIntWriteState	:=	0;
			END_IF
	END_CASE
END_IF




IF bRHskTRG THEN
	CASE nRHskState	OF
		0:
			nRHskBusyIdx	:=	0;
			nRHskState	:=	1;
		1:
			fb_ReadRParams(
				bExecute	:=	TRUE,
				nChnId		:=	inst_NcToPlc_NCI.ChnId,
				pAddr		:=	ADR(nRHskVal),
				nIndex		:=	TO_DINT(UserVar.R_Params[nRHskBusyIdx]),
				nCount		:=	1);
			nRHskState	:=	2;
		2:
			IF fb_ReadRParams.bBusy THEN
				fb_ReadRParams(
					bExecute	:=	FALSE,
					nChnId		:=	inst_NcToPlc_NCI.ChnId,
					pAddr		:=	ADR(nRHskVal),
					nIndex		:=	TO_DINT(UserVar.R_Params[nRHskBusyIdx]),
					nCount		:=	1);
				IF nRHskVal	<>	UserVar.R_InitVal THEN
					fb_ConfirmHsk(
						bExecute	:=	TRUE,
						sNciToPlc	:=	inst_NcToPlc_NCI,
						sPlcToNci	:=	inst_PlcToNc_NCI,);
					nRHskState	:=	3;
				ELSE
					nRHskBusyIdx	:=	nRHskBusyIdx	+	1;
					IF nRHskBusyIdx >=	(SIZEOF(UserVar.R_Params) / 2) THEN
						nRHskState	:=	0;
					ELSE
						nRHskState	:=	1;
					END_IF
				END_IF
			END_IF
		3:
			IF 	fb_ConfirmHsk.bBusy THEN
				fb_ConfirmHsk(
					bExecute	:=	FALSE,
					sNciToPlc	:=	inst_NcToPlc_NCI,
					sPlcToNci	:=	inst_PlcToNc_NCI,);
				bRHskTRG	:=	FALSE;
				nRHskState	:=	0;
			END_IF
	END_CASE
END_IF

END_FUNCTION_BLOCK

// ---- POUs/FB/Keyence/FB_LJ_S8000Capture.TcPOU
FUNCTION_BLOCK FB_LJ_S8000Capture
VAR_INPUT
	bExecute	:	BOOL	:=	FALSE;
END_VAR
VAR_OUTPUT
	bBusy		:	BOOL	:=	FALSE;
END_VAR
VAR
	nState		:	UDINT	:=	0;
END_VAR

CASE nState	OF

0:	
	IF bExecute	THEN
		IF NOT ExtPort.LJ_S8000_bTRG_ack THEN
			ExtPort.LJ_S8000_bTRG	:=	TRUE;
			bBusy	:=	TRUE;
			nState	:=	1;
		END_IF
	END_IF

1:
	IF ExtPort.LJ_S8000_bTRG_ack THEN
		ExtPort.LJ_S8000_bTRG	:=	FALSE;
	END_IF
	IF ExtPort.LJ_S8000_bBusy THEN
		nState	:=	2;
	END_IF
	
2:
	IF ExtPort.LJ_S8000_bReady THEN
		bBusy	:=	FALSE;
		nState	:=	0;
	END_IF
	
END_CASE

END_FUNCTION_BLOCK

// ---- POUs/FB/Nordson/FB_WritePressure.TcPOU
FUNCTION_BLOCK FB_WritePressure
VAR_INPUT
	bExecute	:	BOOL	:=	FALSE;
	Pressure	:	REAL	:=	0.0;
END_VAR
VAR_OUTPUT
	bBusy		:	BOOL	:=	FALSE;
	bErr		:	BOOL	:=	FALSE;
END_VAR
VAR
	nState		:	UDINT	:=	0;
END_VAR

// bNordWriteAcc 키면서 Press 값 넣고
// busy state로 올림

// PYADS에서 press 를 읽어서 입력하고
// 만약 실패시 busy 끄면서 fail 올리고
// 다 입력되면 bNordWriteAcc 끄기


CASE nState OF

0:
	IF bExecute	THEN
		PYADSPort.bNordWriteReq	:=	TRUE;
		PYADSPort.nNordPress	:=	Pressure;
		bBusy	:=	TRUE;
		nState	:=	1;
	END_IF

1:
	IF NOT PYADSPort.bNordWriteReq THEN
		IF PYADSPort.bNordWriteErr THEN
			PYADSPort.bNordWriteErr	:=	FALSE;
			PYADSPort.nNordPress	:=	0.0;
			bErr	:=	TRUE;
		ELSE
			bErr	:=	FALSE;
		END_IF
			bBusy	:=	FALSE;
			nState	:=	0;		
	END_IF
END_CASE

END_FUNCTION_BLOCK

// ---- POUs/FB/MicroFab/FB_PulseInterval.TcPOU
FUNCTION_BLOCK FB_PulseInterval
VAR_INPUT
	bOn			:	BOOL	:=	FALSE;
	nInterval	:	UDINT	:=	100;		// (Rising edge ~ Rising edge, [ms]) Must be multiple of 20
END_VAR
VAR_OUTPUT
END_VAR
VAR
	nClk		:	UDINT	:=	0;
END_VAR

IF	bOn	THEN
	IF nClk	= 0	THEN
		ExtPort.EL2124_OUT[0]	:=	NOT ExtPort.EL2124_OUT[0];
	END_IF
	IF nClk < TO_UDINT(nInterval / (2 * 10)) THEN
		nClk	:=	nClk + 1;
	ELSE		
		nClk	:=	0;
	END_IF
ELSE
	nClk	:=	0;
	ExtPort.EL2124_OUT[0]	:=	FALSE;
END_IF

END_FUNCTION_BLOCK

// ---- POUs/function/f_Contains_INT.TcPOU
FUNCTION f_Contains_INT : BOOL
VAR_INPUT
    num	: INT;
END_VAR
VAR_IN_OUT
	arr : ARRAY[*] OF INT;   // 가변 길이 1D 배열
END_VAR
VAR
    i : DINT;
END_VAR

F_Contains_INT := FALSE;

FOR i := LOWER_BOUND(arr, 1) TO UPPER_BOUND(arr, 1) DO
    IF arr[i] = num THEN
        F_Contains_INT := TRUE;
        RETURN;
    END_IF
END_FOR

END_FUNCTION

// ---- POUs/FB/FB_RParamInit.TcPOU
FUNCTION_BLOCK FB_RParamInit
VAR_INPUT
	bExecute	:	BOOL	:=	FALSE;
END_VAR
VAR_OUTPUT
	bBusy		:	BOOL	:=	FALSE;
	bErr		:	BOOL	:=	FALSE;
END_VAR
VAR_IN_OUT
	inst_NcToPlc_NCI	:	NCTOPLC_NCICHANNEL_REF;
END_VAR
VAR
	BusyIdx		:	DINT	:=	0;	
	nState		:	DINT	:=	0;
	fb_WriteRParams	:	ItpWriteRParams;
END_VAR

CASE nState OF
	
0:
	IF bExecute THEN
		bBusy	:=	TRUE;
		bErr	:=	FALSE;
		nState	:=	1;
		BusyIdx	:=	0;
	END_IF

1:
	fb_WriteRParams(
		bExecute	:=	TRUE,
		nChnId		:=	inst_NcToPlc_NCI.ChnId,
		pAddr		:=	ADR(UserVar.R_InitVal),
		nIndex		:=	TO_DINT(UserVar.R_Params[BusyIdx]),
		nCount		:=	1);
	nState	:=	2;


2:
	IF fb_WriteRParams.bBusy THEN
		fb_WriteRParams(
			bExecute	:=	FALSE,
			nChnId		:=	inst_NcToPlc_NCI.ChnId,
			pAddr		:=	ADR(UserVar.R_InitVal),
			nIndex		:=	TO_DINT(UserVar.R_Params[BusyIdx]),
			nCount		:=	1);
		nState	:=	3;
	END_IF
	

3:	
	fb_WriteRParams(	bExecute	:=	FALSE);
	IF NOT fb_WriteRParams.bBusy THEN
		IF fb_WriteRParams.bErr THEN
			bErr	:=	TRUE;
			bBusy	:=	FALSE;
			nState	:=	0;
		ELSE
			BusyIdx	:=	BusyIdx	+	1;
			IF BusyIdx 	>=	(SIZEOF(UserVar.R_Params) / 2) THEN
				bBusy	:=	FALSE;
				nState	:=	0;
			ELSE
				nState	:=	1;
			END_IF
		END_IF
	END_IF

END_CASE

END_FUNCTION_BLOCK

// ---- POUs/FB/FB_BackendManager.TcPOU
FUNCTION_BLOCK FB_BackendManager
VAR_INPUT
END_VAR
VAR_OUTPUT
END_VAR
VAR
	BackendStartState	:	UDINT	:=	0;
	
	fbStart  : NT_StartProcess;
	fb_TimeCalc	:	FB_TimeCalculator;
	bTimerActive	:	BOOL	:=	FALSE;
	nTimerState	:	UDINT	:=	0;
	nTimerCnt	:	UDINT	:=	0;
END_VAR

CASE BackendStartState OF
	0:
		fbStart(
			NETID     := '',
			PATHSTR   := 'C:\ProgramData\miniconda3\envs\ERC_CONTROL_BACKEND\pythonw.exe',
			DIRNAME   := 'C:\Users\Administrator\Documents\ERC\PythonProjects\PythonBackend\NCI_260109',
			COMNDLINE := '"C:\Users\Administrator\Documents\ERC\PythonProjects\PythonBackend\NCI_260109\main.py"',
			START     := TRUE,
			TMOUT     := T#5S
		);
		IF fbStart.BUSY THEN
			BackendStartState	:=	1;
		END_IF
	
	1:
		fbStart(START:=	FALSE);
		BackendStartState	:=	2;
		UserVar.bBackendStarted	:=	TRUE;
		PYADSPort.bHeartbeat	:=	TRUE;
		bTimerActive	:=	TRUE;
		
	2:
		IF nTimerCnt >= 200 THEN
			BackendStartState	:=	3;
			nTimerCnt	:=	0;
		END_IF
	
	3:
		IF nTimerCnt >= 50 THEN
			PYADSPort.bHeartbeat	:=	TRUE;
			BackendStartState	:=	4;
		END_IF
	4:
		IF nTimerCnt >= 100 THEN
			IF UserVar.gInSync THEN
				nTimerCnt	:=	0;
				BackendStartState	:=	3;
			ELSE
				UserVar.bBackendStarted	:=	FALSE;
				bTimerActive	:=	FALSE;
				nTimerCnt	:=	0;
				BackendStartState	:=	0;
			END_IF
		END_IF
		
END_CASE


IF bTimerActive	THEN
	fb_TimeCalc();
	nTimerCnt	:=	nTimerCnt + 1;
END_IF

END_FUNCTION_BLOCK

// ---- POUs/FB/FB_TimeCalculator.TcPOU
FUNCTION_BLOCK FB_TimeCalculator
VAR
	fbLocalTime		:	FB_LocalSystemTime := (bEnable := TRUE, dwCycle := 1);

    stPy      : TIMESTRUCT;
	
	
	    // 추가: Timezone 정보 & 변환 FB
    fbGetTz   : FB_GetTimeZoneInformation;
    fbLoc2Utc : FB_TzSpecificLocalTimeToSystemTime;
    fbUtc2Loc : FB_SystemTimeToTzSpecificLocalTime;

    tzInfo    : ST_TimeZoneInformation;
    bTzReady  : BOOL := FALSE;

    stNowLocal : TIMESTRUCT;
    stNowUtc   : TIMESTRUCT;

    dtNowUtc   : DT;
    dtPy       : DT;

    nowSec     : DWORD;
    pySec      : DWORD;
    diff       : LINT;

    stPyUtc    : TIMESTRUCT;
    stPyLocal  : TIMESTRUCT;
END_VAR

// 0) Timezone 정보 1회 확보 (부팅 후 한 번만)
IF NOT bTzReady THEN
    fbGetTz(bExecute := TRUE, sNetID := '');
    IF (NOT fbGetTz.bBusy) THEN
        IF (NOT fbGetTz.bError) THEN
            tzInfo   := fbGetTz.tzInfo;
            bTzReady := TRUE;
        END_IF
    END_IF
END_IF

// 1) 로컬 시간 업데이트
fbLocalTime();

IF bTzReady AND fbLocalTime.bValid THEN
    // (A) PLC 로컬(Seoul) 시간
    stNowLocal := fbLocalTime.systemTime;

    // (B) 로컬 -> UTC 변환 후 DT로 변환 (비교 기준 통일)
    fbLoc2Utc(in := stNowLocal, tzInfo := tzInfo, out => stNowUtc);
    stNowUtc.wMilliseconds := 0;
    dtNowUtc := SYSTEMTIME_TO_DT(stNowUtc);

    // (C) Python에서 받은 DT (권장: UTC epoch seconds로 write됨)
    dtPy := PYADSPort.dtHeartbeatTime;

    // (D) 초 단위 비교
    nowSec := DT_TO_DWORD(dtNowUtc);
    pySec  := DT_TO_DWORD(dtPy);
    diff   := DWORD_TO_LINT(nowSec) - DWORD_TO_LINT(pySec);

    UserVar.gDiffSec := diff;
    UserVar.gInSync  := (ABS(diff) <= 5);

    // (E) 표시용 문자열
    // PLC 로컬(Seoul) 표시
    UserVar.gPlcStr := SYSTEMTIME_TO_STRING(stNowLocal);

    // Python(UTC DT) -> 로컬(Seoul)로 변환해서 표시
    stPyUtc := DT_TO_SYSTEMTIME(dtPy);
    fbUtc2Loc(in := stPyUtc, tzInfo := tzInfo, out => stPyLocal);
    UserVar.gPyStr := SYSTEMTIME_TO_STRING(stPyLocal);
END_IF

END_FUNCTION_BLOCK

// ---- POUs/FB/FB_Jog.TcPOU
FUNCTION_BLOCK FB_Jog
VAR_INPUT
	JogButton	:	INT;
END_VAR
VAR_OUTPUT
	bBusy		:	BOOL;
	bError		:	BOOL;
END_VAR
VAR_IN_OUT
	mot			:	AXIS_REF;
END_VAR
VAR
	fb_MCJog	:	MC_Jog;
END_VAR

CASE ABS(JogButton) OF
	0:	fb_MCJog(
			Axis	:=	mot);
	1:	fb_MCJog(
			Axis	:=	mot,
			Mode	:=	E_JogMode.MC_JOGMODE_STANDARD_SLOW);
	2:	fb_MCJog(
			Axis	:=	mot,
			Mode	:=	E_JogMode.MC_JOGMODE_STANDARD_FAST);
	3:	fb_MCJog(
			Axis	:=	mot,
			Mode	:=	E_JogMode.MC_JOGMODE_CONTINOUS,
			Velocity:=	STRING_TO_LREAL(UserVar.JogTargVel)/60.0);
END_CASE

IF JogButton > 0 THEN
	fb_MCJog.JogForward	:=	TRUE;
	fb_MCJog.JogBackwards	:=	FALSE;
END_IF

IF JogButton < 0 THEN
	fb_MCJog.JogForward	:=	FALSE;
	fb_MCJog.JogBackwards	:=	TRUE;
END_IF

IF JogButton = 0 THEN
	fb_MCJog.JogForward	:=	FALSE;
	fb_MCJog.JogBackwards	:=	FALSE;
END_IF

bBusy	:=	fb_MCJog.Busy;
bError	:=	fb_MCJog.Error;

END_FUNCTION_BLOCK

// ---- POUs/FB/FB_ExtMessage.TcPOU
FUNCTION_BLOCK FB_ExtMessage
VAR_INPUT
END_VAR
VAR_OUTPUT

	
END_VAR
VAR_IN_OUT
	motX:	AXIS_REF;
	motY:	AXIS_REF;
	motZ:	AXIS_REF;
	bBusy	:	BOOL;
	inst_NcToPlc_NCI	:	NCTOPLC_NCICHANNEL_REF;
	inst_PlcToNc_NCI	:	PLCTONC_NCICHANNEL_REF;
END_VAR

VAR
	ActPosX	:	LREAL;
	ActPosY	:	LREAL;
	ActPosZ	:	LREAL;
	
	ActVelX	:	LREAL;
	ActVelY	:	LREAL;
	ActVelZ	:	LREAL;
	
	ActAccX	:	LREAL;
	ActAccY	:	LREAL;
	ActAccZ	:	LREAL;
	
	SetPosX	:	LREAL;
	SetPosY	:	LREAL;
	SetPosZ	:	LREAL;
	
	SetVelX	:	LREAL;
	SetVelY	:	LREAL;
	SetVelZ	:	LREAL;
	
	SetAccX	:	LREAL;
	SetAccY	:	LREAL;
	SetAccZ	:	LREAL;


	fb_AdsRead	:	ADSREAD;
	nTimerCnt	:	UDINT	:=	0;
END_VAR

ActPosX	:=	motX.NcToPlc.ActPos;
ActPosY	:=	motY.NcToPlc.ActPos;
ActPosZ	:=	motZ.NcToPlc.ActPos;

ActVelX	:=	motX.NcToPlc.ActVelo;
ActVelY	:=	motY.NcToPlc.ActVelo;
ActVelZ	:=	motZ.NcToPlc.ActVelo;

ActAccX	:=	motX.NcToPlc.ActAcc;
ActAccY	:=	motY.NcToPlc.ActAcc;
ActAccZ	:=	motZ.NcToPlc.ActAcc;

SetPosX	:=	motX.NcToPlc.SetPos;
SetPosY	:=	motY.NcToPlc.SetPos;
SetPosZ	:=	motZ.NcToPlc.SetPos;

SetVelX	:=	motX.NcToPlc.SetVelo;
SetVelY	:=	motY.NcToPlc.SetVelo;
SetVelZ	:=	motZ.NcToPlc.SetVelo;

SetAccX	:=	motX.NcToPlc.SetAcc;
SetAccY	:=	motY.NcToPlc.SetAcc;
SetAccZ	:=	motZ.NcToPlc.SetAcc;

HMIVar.sActPosX  :=  LREAL_TO_FMTSTR(ActPosX, 3, TRUE);
HMIVar.sActPosY  :=  LREAL_TO_FMTSTR(ActPosY, 3, TRUE);
HMIVar.sActPosZ  :=  LREAL_TO_FMTSTR(ActPosZ, 3, TRUE);

HMIVar.sActVelX  :=  LREAL_TO_FMTSTR(ActVelX, 3, TRUE);
HMIVar.sActVelY  :=  LREAL_TO_FMTSTR(ActVelY, 3, TRUE);
HMIVar.sActVelZ  :=  LREAL_TO_FMTSTR(ActVelZ, 3, TRUE);

HMIVar.sActAccX  :=  LREAL_TO_FMTSTR(ActAccX, 3, TRUE);
HMIVar.sActAccY  :=  LREAL_TO_FMTSTR(ActAccY, 3, TRUE);
HMIVar.sActAccZ  :=  LREAL_TO_FMTSTR(ActAccZ, 3, TRUE);

HMIVar.sSetPosX  :=  LREAL_TO_FMTSTR(SetPosX, 3, TRUE);
HMIVar.sSetPosY  :=  LREAL_TO_FMTSTR(SetPosY, 3, TRUE);
HMIVar.sSetPosZ  :=  LREAL_TO_FMTSTR(SetPosZ, 3, TRUE);

HMIVar.sSetVelX  :=  LREAL_TO_FMTSTR(SetVelX, 3, TRUE);
HMIVar.sSetVelY  :=  LREAL_TO_FMTSTR(SetVelY, 3, TRUE);
HMIVar.sSetVelZ  :=  LREAL_TO_FMTSTR(SetVelZ, 3, TRUE);

HMIVar.sSetAccX  :=  LREAL_TO_FMTSTR(SetAccX, 3, TRUE);
HMIVar.sSetAccY  :=  LREAL_TO_FMTSTR(SetAccY, 3, TRUE);
HMIVar.sSetAccZ  :=  LREAL_TO_FMTSTR(SetAccZ, 3, TRUE);

HMIVar.EstimatedTime	:=	CONCAT(LREAL_TO_FMTSTR(PYADSPort.nEstTime, 3, TRUE), 's');



HMIVar.bNaviActive	:=	(NOT bBusy);

IF (UserVar.Auto_CodeType <> 0) THEN
	IF  HMIVar.CodeName <> '' THEN
		CASE UserVar.Auto_CodeType OF
		1:
			IF f_QueuePush(HMIVar.CodeName, ADR(UserVar.GCodeNameQueue)) THEN
				UserVar.Auto_CodeType	:=	0;
				HMIVar.GCodeQueueString	:=	f_Queue_ToString(ADR(UserVar.GCodeNameQueue));
			END_IF
//			UserVar.QueuedGCodeName	:=	HMIVar.CodeName;	
		END_CASE		
	ELSE
		UserVar.Auto_CodeType	:=	0;
	END_IF
	
END_IF



UserVar.CurrBlockNum	:=	ItpGetBlockNumber(inst_NcToPlc_NCI);

IF UserVar.CurrBlockNum <> 0 THEN
	HMIVar.CurrBlockNumSTR	:=	CONCAT('N', UDINT_TO_STRING(UserVar.CurrBlockNum));
ELSE
	HMIVar.CurrBlockNumSTR	:=	'-';
END_IF

END_FUNCTION_BLOCK

// ---- POUs/function/f_QueuePush.TcPOU
FUNCTION f_QueuePush : BOOL
VAR_INPUT
    str : STRING(255);
    pQueue : POINTER TO T_StringQueue;
END_VAR
VAR
END_VAR

IF pQueue^.Count >= 20 THEN
    f_QueuePush := FALSE; // Full
ELSE
    pQueue^.Buffer[pQueue^.Tail] := str;
    pQueue^.Tail := (pQueue^.Tail + 1) MOD 20;
    pQueue^.Count := pQueue^.Count + 1;
    f_QueuePush := TRUE;
END_IF

END_FUNCTION

// ---- POUs/function/f_Queue_ToString.TcPOU
FUNCTION f_Queue_ToString : STRING(8192)
VAR_INPUT
    pQueue : POINTER TO T_StringQueue;
END_VAR
VAR
    i       : INT;
    idx     : INT;
    result  : STRING(8192);
    tmp     : STRING(255);
END_VAR

result := '';
idx := pQueue^.Head;

FOR i := 1 TO pQueue^.Count DO
    tmp := pQueue^.Buffer[idx];

    // 내용 추가
//    result := CONCAT(result, tmp);
	CONCAT2(
        pSrcString1 := ADR(result),
        pSrcString2 := ADR(tmp),
        pDstString  := ADR(result),
        nDstSize    := SIZEOF(result)
    );

    // 마지막 요소가 아니면 엔터 추가
    IF i < pQueue^.Count THEN
//        result := CONCAT(result, '\r\n');
        CONCAT2(
            pSrcString1 := ADR(result),
            pSrcString2 := ADR('$R$N'),
            pDstString  := ADR(result),
            nDstSize    := SIZEOF(result)
        );
    END_IF

    // 원형 인덱스 이동
    idx := (idx + 1) MOD 20;
END_FOR

f_Queue_ToString := result;

END_FUNCTION

// ---- POUs/FB/FB_HMITask.TcPOU
FUNCTION_BLOCK FB_HMITask
VAR_INPUT
END_VAR
VAR_OUTPUT
END_VAR
VAR
	fb_ReadPres					:	FB_ReadPressure;
	fb_WritePres				:	FB_WritePressure;
	fb_LJ_S8000Cap				:	FB_LJ_S8000Capture;
	
	nNordsonReadPressureCase	:	UDINT	:=	0;
	nNordsonWritePressureCase	:	UDINT	:=	0;
	nLJ_S8000CaptureCase		:	UDINT	:=	0;
	
	nClearQueueCase				:	UDINT	:=	0;
END_VAR

      IF UserVar.NordsonReadPressureBtn	THEN
	CASE nNordsonReadPressureCase OF
		0:
			UserVar.NordsonPressureActive	:=	FALSE;
			fb_ReadPres( bExecute	:=	TRUE);
			IF fb_ReadPres.bBusy	THEN
				fb_ReadPres.bExecute	:=	FALSE;
				nNordsonReadPressureCase	:=	1;
			END_IF
		1:
			fb_ReadPres( bExecute	:=	FALSE);
			IF NOT fb_ReadPres.bBusy THEN
				IF NOT fb_ReadPres.bErr THEN
					HMIVar.NordsonPressure	:=	REAL_TO_STRING(fb_ReadPres.Pressure);
				ELSE
					HMIVar.NordsonPressure	:=	'0';
				END_IF
				UserVar.NordsonPressureActive	:=	TRUE;
				UserVar.NordsonReadPressureBtn	:=	FALSE;
				nNordsonReadPressureCase	:=	0;
			END_IF
	END_CASE
END_IF


IF UserVar.NordsonWritePressureBtn	THEN
	CASE nNordsonWritePressureCase OF
		0:
			UserVar.NordsonPressureActive	:=	FALSE;
			fb_WritePres(
				bExecute	:=	TRUE,
				Pressure	:=	STRING_TO_REAL(HMIVar.NordsonPressure));
			IF fb_WritePres.bBusy	THEN
				fb_WritePres.bExecute	:=	FALSE;
				nNordsonWritePressureCase	:=	1;
			END_IF
		1:
			fb_WritePres(
				bExecute	:=	FALSE);
			IF NOT fb_WritePres.bBusy THEN
				UserVar.NordsonPressureActive	:=	TRUE;
				UserVar.NordsonWritePressureBtn	:=	FALSE;
				nNordsonWritePressureCase	:=	0;
			END_IF
	END_CASE
END_IF


IF UserVar.LJ_S8000CaptureBtn	THEN
	CASE nLJ_S8000CaptureCase OF
		0:
			UserVar.LJ_S8000CaptureActive	:=	FALSE;
			fb_LJ_S8000Cap(	bExecute :=	TRUE);
			IF fb_LJ_S8000Cap.bBusy THEN
				fb_LJ_S8000Cap.bExecute	:=	FALSE;
				nLJ_S8000CaptureCase	:=	1;
			END_IF
		1:
			fb_LJ_S8000Cap(	bExecute :=	FALSE);
			IF NOT fb_LJ_S8000Cap.bBusy THEN
				UserVar.LJ_S8000CaptureActive	:=	TRUE;
				UserVar.LJ_S8000CaptureBtn	:=	FALSE;
				nLJ_S8000CaptureCase	:=	0;
			END_IF
	END_CASE
END_IF


IF UserVar.bClearQueue THEN	
	CASE nClearQueueCase OF
		0:
			IF NOT f_QueuePop(pQueue := ADR(UserVar.GCodeNameQueue)) THEN
				nClearQueueCase	:=	1;
			END_IF
		1:
			HMIVar.GCodeQueueString	:=	f_Queue_ToString(ADR(UserVar.GCodeNameQueue));
			UserVar.bClearQueue	:=	FALSE;
			nClearQueueCase	:=	0;
	END_CASE
END_IF



IF ExtPort.EL1008_IN[1] THEN
	UserVar.bNordsonFoot	:=	 TRUE;
	ExtPort.EL2634_OUT[0]	:=	TRUE;
END_IF


IF UserVar.bNordsonFoot	THEN
	IF NOT ExtPort.EL1008_IN[1]	THEN
		UserVar.bNordsonFoot	:=	FALSE;
		ExtPort.EL2634_OUT[0]	:=	FALSE;
	END_IF
END_IF

END_FUNCTION_BLOCK

// ---- POUs/FB/Nordson/FB_ReadPressure.TcPOU
FUNCTION_BLOCK FB_ReadPressure
VAR_INPUT
	bExecute	:	BOOL	:=	FALSE;
END_VAR
VAR_OUTPUT
	bBusy		:	BOOL	:=	FALSE;
	bErr		:	BOOL	:=	FALSE;
	Pressure	:	REAL	:=	0.0;
END_VAR
VAR
	nState		:	UDINT	:=	0;
END_VAR

// bNordReadAcc 키면서
// busy state로 올림

// press 읽어서 PYADS에 입력하고
// 다 입력되면 NordPress에 쓰고 bNordReadAcc 끄기
// 만약 실패시 busy 끄면서 fail 올리기



CASE nState OF

0:
	IF bExecute	THEN
		PYADSPort.bNordReadReq	:=	TRUE;
		bBusy	:=	TRUE;
		nState	:=	1;
	END_IF

1:
	IF NOT PYADSPort.bNordReadReq THEN
		IF PYADSPort.bNordReadErr THEN
			PYADSPort.bNordReadErr	:=	FALSE;
			bErr	:=	TRUE;
		ELSE
			bErr	:=	FALSE;
		END_IF
			Pressure:=	PYADSPort.nNordPress;
			bBusy	:=	FALSE;
			nState	:=	0;
	END_IF
END_CASE

END_FUNCTION_BLOCK

// ---- POUs/function/f_QueuePop.TcPOU
FUNCTION f_QueuePop : BOOL
VAR_INPUT
    pQueue : POINTER TO T_StringQueue;
END_VAR
VAR_OUTPUT
    str : STRING(255);
END_VAR

IF pQueue^.Count <= 0 THEN
    f_QueuePop := FALSE; // Empty
ELSE
    str := pQueue^.Buffer[pQueue^.Head];
    pQueue^.Head := (pQueue^.Head + 1) MOD 20;
    pQueue^.Count := pQueue^.Count - 1;
    f_QueuePop := TRUE;
END_IF

END_FUNCTION

// ---- POUs/function/f_MakeAbsPath.TcPOU
FUNCTION f_MakeAbsPath : STRING(255)
VAR_INPUT
	GCodePath	:	STRING(255);
END_VAR
VAR
END_VAR

f_MakeAbsPath	:=	CONCAT(UserVar.GCodeBasePath, GCodePath);

END_FUNCTION
